Fanuc KAREL source: KT00600.KL

PROGRAM KT00600
%NOLOCKGROUP
VAR
  I1: INTEGER
  I2: INTEGER
  OUT: BOOLEAN
BEGIN
  I1 = 2
  I2 = 3
  I1 = 2
  I2 = 3
  OUT = NOT I1
END KT00600
